Fanuc KAREL source: kb00094.KL

-- PROVISIONAL review KL for V770-1; original PC SHA256 def808471585a7b8c8160940bd6c6735b8123c7c3f8c3f4e994c7820a729c394
-- Incomplete behavior may be omitted. Consult companion uncertainty JSON. Do not deploy.
PROGRAM KB00094
%NOLOCKGROUP
BEGIN
  -- UNRESOLVED_PC offsets 5-12; opcodes 9D,23
  -- UNRESOLVED_PC offsets 17-27; opcodes 27,22,31
  -- UNRESOLVED_PC offsets 32-36; opcodes 7F
END KB00094
